{region 'Documentation'}
(*!
<summary>Checks equality with the expected UINT value.</summary>
*)
{endregion}
FUNCTION_BLOCK AssertEqual_UInt EXTENDS AssertionBase
VAR_INPUT
    IN : UINT; //! Actual value checked or observed by this Assertion.
    Expected : UINT; //! Reference value for comparison with IN.
END_VAR

SUPER^();

{region 'Documentation'}
(*!
<summary>Check equality with the expected UINT value.</summary>
*)
{endregion}
METHOD PROTECTED Assert
VAR
    Message : STRING(GVL_Constants.MessageLength);
    ExpectedText : STRING(GVL_Constants.AssertionValueLength);
    ActualText : STRING(GVL_Constants.AssertionValueLength);
END_VAR
IF NOT EvaluationActive THEN
    RETURN;
END_IF;

IF Result = E_Result.Error THEN
    RETURN;
END_IF;

IF Result = E_Result.Failed THEN
    RETURN;
END_IF;

IF IN <> Expected THEN
    ExpectedText := UINT_TO_STRING(Expected);
    ActualText := UINT_TO_STRING(IN);
    Message := CONCAT('Assertion failed: values are not equal. Expected = ',
        ExpectedText);
    Message := CONCAT(Message, ', Actual = ');
    Message := CONCAT(Message, ActualText);
    Message := CONCAT(Message, '.');
    Fail(Message := Message);
    RETURN;
END_IF;

Pass();
END_METHOD

END_FUNCTION_BLOCK

(* stored: Version 1.1.0.1
   POU AssertEqual_UInt: Id {ab32cad3-9c6b-444e-b9d1-290228020346}, SpecialFunc None
   Folder Internal: Id {76098aad-b7b9-4e3a-be1f-ee2d0dff59ee}
   Method Assert: Id {99972bef-0cda-4ac7-bd8d-bfac39b09bd4} *)
